// TIA Portal V21 export
VAR_GLOBAL   // PLC tag table "IO_Einschubachse"
   ModePos_z AT %MW4 : Int;
   AxisRef_z AT %M6.0 : Bool;
   Error_z AT %M13.0 : Bool;
   ActVel_z AT %M60.0 : LReal;
   ActPos_z AT %M80.0 : LReal;
   AxisEnabled_z AT %M13.1 : Bool;
   ErrorID_z AT %MW90 : Word;
END_VAR
